// TIA Portal V21 export
// export: Created 2026-11-21T13:24:04.2913446Z, ExportSetting WithDefaults, DisplayName Totally Integrated Automation Portal, DisplayVersion V21, DisplayName STEP 7 Professional, DisplayVersion V21, DisplayName STEP 7 Safety, DisplayVersion V21, DisplayName Tech WebApplication, DisplayVersion V21, DisplayName WinCC Basic/Comfort/Advanced, DisplayVersion V21, DisplayName WinCC Unified, DisplayVersion V21
FUNCTION "Enable" : Bool   // FC2, F_LAD
{ S7_Optimized_Access := 'TRUE' }
VERSION : 0.1
// True while both inputs are true.
// stored: AutoNumber true, IsIECCheckEnabled false, UDAEnableTagReadback false
   VAR_INPUT
      "a" : Bool;
      "b" : Bool;
   END_VAR
BEGIN

REGION Network 1: Both inputs
   // On while both inputs are on.
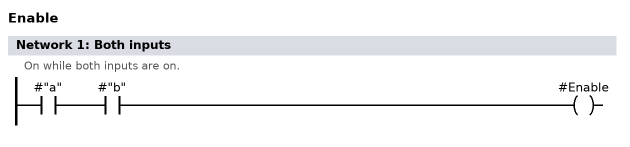
   RUNG wire#powerrail
      Contact( #"a" )
      Contact( #"b" )
      Coil( #Enable )
   END_RUNG
   // the same network as SCL:
   #Enable := #"a" AND #"b";
END_REGION
END_FUNCTION
